TYPE ST_PolarIIChamber_Recipe :
STRUCT
	AcidDropOffset : LREAL; // deg
	StrokePositiveLimit : LREAL; // deg
	StrokeNegativeLimit : LREAL; // deg
	SpeedAtPosition : ARRAY[1..50] OF LREAL; // RPM, from negative to positive limit
END_STRUCT
END_TYPE

(* stored: Version 1.1.0.1, ProductVersion 3.1.4026.18
   DUT ST_PolarIIChamber_Recipe: Id {14000000-0000-0000-0000-000000000008} *)
